// TIA Portal V21 export
// export: Created 2026-11-07T15:50:59.9946565Z, ExportSetting WithDefaults, DisplayName Totally Integrated Automation Portal, DisplayVersion V21, DisplayName STEP 7 Professional, DisplayVersion V21, DisplayName STEP 7 Safety, DisplayVersion V21, DisplayName Tech WebApplication, DisplayVersion V21, DisplayName WinCC Basic/Comfort/Advanced, DisplayVersion V21, DisplayName WinCC Unified, DisplayVersion V21
TextList "TL_Order"  ListRange=Decimal
  TextListEntry   EntryType=SingleValue, Text="0 slobodan redoslijed"
  TextListEntry   EntryType=SingleValue, From=1, To=1, Text="1 redoslijed po listi"
  TextListEntry   EntryType=SingleValue, From=2, To=2, Text="2 strogo: istovar pa ukrcaj"
